(* PLC project Vn_op_sin, Beckhoff Automation GmbH TwinCAT PLC Control 3.5.13.21 *)
(* stored: creationDateTime 1970-01-01T00:00:00 *)

PROGRAM Vn_op_sin

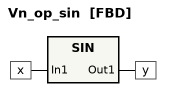
(* FBD diagram, written out as Structured Text *)
y := SIN(x);
END_PROGRAM
